(* IEC 61131-3 sources: ZPLC/packages/zplc-ide/plant-scenes/counted-queue, 2 files *)

(* ---- reference.st ---- *)
PROGRAM CountedQueue
VAR_INPUT
    Start  AT %I0.0 : BOOL;
    EyeIn  AT %I0.1 : BOOL;
    EyeOut AT %I0.2 : BOOL;
END_VAR
VAR_OUTPUT
    Run  AT %Q0.0 : BOOL;
    Emit AT %Q0.1 : BOOL;
    Done AT %Q0.2 : BOOL;
END_VAR
VAR
    Active   : BOOL;
    Loaded   : CTU;
    Unloaded : CTU;
    InGone   : F_TRIG;
END_VAR

IF Start THEN
    Active := TRUE;
END_IF;

Loaded(CU := EyeIn, R := FALSE, PV := 3);
Unloaded(CU := EyeOut, R := FALSE, PV := 3);
InGone(CLK := EyeIn);

(* the first box on Start, each next box once the previous one has left the emitter *)
Emit := (Start OR InGone.Q) AND Active AND NOT Loaded.Q;
Done := Unloaded.Q;
Run := Active AND NOT Unloaded.Q;

END_PROGRAM

(* ---- starter.st ---- *)
PROGRAM CountedQueue
VAR_INPUT
    Start  AT %I0.0 : BOOL;  (* StartButton.pressed: start the batch *)
    EyeIn  AT %I0.1 : BOOL;  (* EyeIn.detect: sees each box that has been loaded *)
    EyeOut AT %I0.2 : BOOL;  (* EyeOut.detect: sees each box about to be unloaded *)
END_VAR
VAR_OUTPUT
    Run  AT %Q0.0 : BOOL;    (* Belt1.run: run the belt *)
    Emit AT %Q0.1 : BOOL;    (* Emitter1.emit: put one box on the belt *)
    Done AT %Q0.2 : BOOL;    (* DoneLight.lit: lit when the batch is finished *)
END_VAR

(* Goal: a press of the start button loads three boxes, one at a time, and
   counts them at EyeIn; then the belt unloads them and a second counter at
   EyeOut tells when all three are gone. Light Done at the end. *)

END_PROGRAM
